Fanuc KAREL source: KA00189.KL

PROGRAM KA00189
%NOLOCKGROUP
VAR
  SRC: ARRAY[4] OF BYTE
  DST: ARRAY[4] OF JOINTPOS
BEGIN
  DST = SRC
END KA00189
